// Riceve i comandi dell'HMI con numero di sequenza (Hmi.Cmd): bNew vale TRUE per un ciclo quando arriva un
// comando nuovo; chi lo esegue risponde con Ack(). nAck/eResult vanno in Hmi.Sts.
// Al primo ciclo dopo l'avvio del PLC il comando presente non si esegue (si allinea nAck): niente comandi
// vecchi rieseguiti dopo un riavvio.
FUNCTION_BLOCK FB_HmiCommandHandler
VAR_INPUT
	stCmd			: ST_HmiCmd;
END_VAR
VAR_OUTPUT
	bNew			: BOOL;
	nAck			: UDINT;
	eResult			: E_HmiResult;
END_VAR
VAR
	bInit			: BOOL;
END_VAR

IF NOT bInit THEN
	bInit := TRUE;
	nAck := stCmd.nSeq;
END_IF

bNew := stCmd.nSeq <> nAck AND stCmd.eCommand <> E_HmiCommand.None;
IF stCmd.nSeq <> nAck AND stCmd.eCommand = E_HmiCommand.None THEN
	nAck := stCmd.nSeq;
	eResult := E_HmiResult.UnknownCommand;
END_IF

// Risposta al comando nuovo di questo ciclo.
METHOD Ack
VAR_INPUT
	eAnswer		: E_HmiResult;
END_VAR
nAck := stCmd.nSeq;
eResult := eAnswer;
bNew := FALSE;
END_METHOD

END_FUNCTION_BLOCK

(* stored: Version 1.1.0.1, ProductVersion 3.1.4024.12
   POU FB_HmiCommandHandler: Id {5f32afa4-72c2-4fa2-b180-ae8929bf1bba}, SpecialFunc None
   Method Ack: Id {278b14c6-a18b-460d-9c1b-c13387ba0d7f} *)
